SUBAPPLICATION NetEv_Einmal (* Event nur beim ersten Mal durchlassen, danach EO1 *)
  (* Standard: 61499-2; Description: Copyright (c) 2026 Meisterschulen am Ostbahnhof This program and the accompanying materials are made available under the terms of the Eclipse Public License 2.0 which is available at https://www.eclipse.org/legal/epl-2.0/ SPDX-License-Identifier: EPL-2.0 *)
  (* Version 1.0, 2026-11-17, Franz Höpfinger, Meisterschulen am Ostbahnhof, initial implementation *)
  PACKAGE MyLib::sys;
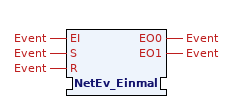
  EVENT_INPUT
    EI; (* Anforderung *)
    S; (* erledigt, ab jetzt EO1 *)
    R; (* zurücksetzen, wieder EO0 *)
  END_EVENT
  EVENT_OUTPUT
    EO0; (* erstes Mal *)
    EO1; (* schon erledigt *)
  END_EVENT
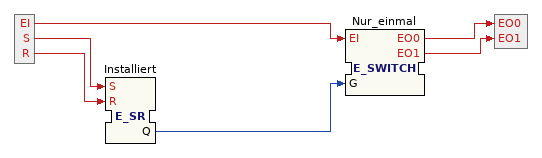
  FBS
    Nur_einmal : iec61499::events::E_SWITCH;
    Installiert : iec61499::events::E_SR;
  END_FBS
  EVENT_CONNECTIONS
    EI TO Nur_einmal.EI;
    S TO Installiert.S;
    R TO Installiert.R;
    Nur_einmal.EO0 TO EO0;
    Nur_einmal.EO1 TO EO1;
  END_CONNECTIONS
  DATA_CONNECTIONS
    Installiert.Q TO Nur_einmal.G;
  END_CONNECTIONS
END_SUBAPPLICATION
